(* PLC project POC, CODESYS CODESYS V3.5 SP22 Patch 4 *)
(* stored: creationDateTime 2026-11-11T00:00:00, modificationDateTime 2026-11-11T00:00:00 *)

PROGRAM PLC_PRG
  VAR
    BT_TESTE : BOOL;
    FALHA_TESTE : BOOL;
    EST_TESTE : BOOL;
  END_VAR

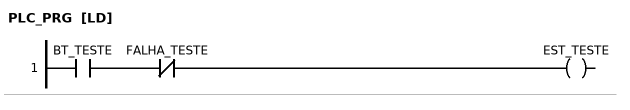
(* LD diagram, written out as Structured Text *)
EST_TESTE := BT_TESTE AND NOT FALHA_TESTE;
END_PROGRAM
